Fanuc KAREL source: KT00352.KL

PROGRAM KT00352
%NOLOCKGROUP
VAR
  P1: XYZWPR
  P2: XYZWPR
  OUT: BOOLEAN
BEGIN
  P1.X = 1.0
  P2.Y = 2.0
  P1.X = 1.0
  P2.Y = 2.0
  OUT = P1 < P2
END KT00352
